FUNCTION_BLOCK basicUVTrojan (* Logica do sistema UV Trojan UV3000Plus (monitoracao Modbus TCP) *)
  (* Standard: 61499-2 *)
  (* Version 1.0, 19/10/2026, Hidryco, Hidryco, 1.0: leitura 41001-41008, canais 1 e 2 (41021-41037, 41061-41077), limpeza 41181-41191; heartbeat 40006 b1 e vigia do heartbeat do SCC *)
  PACKAGE Hidryco.HidrycoLib;
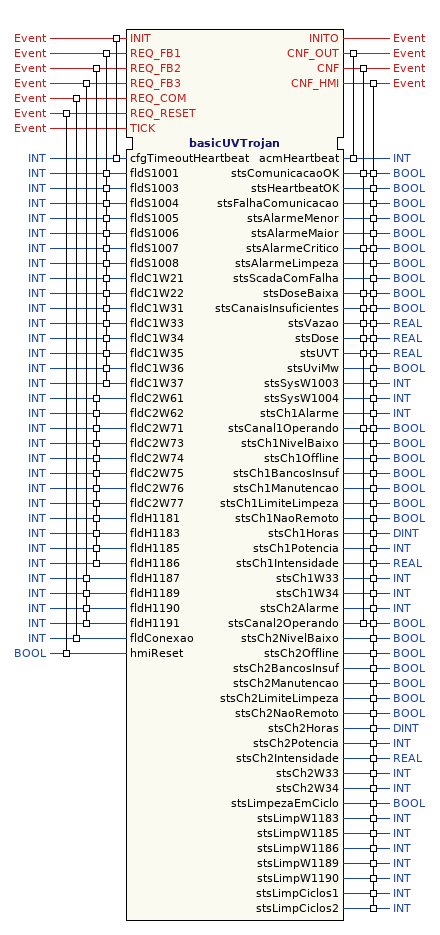
  EVENT_INPUT
    INIT WITH cfgTimeoutHeartbeat; (* Inicializacao *)
    REQ_FB1 WITH fldS1001, fldS1003, fldS1004, fldS1005, fldS1006, fldS1007, fldS1008, fldC1W21, fldC1W22, fldC1W31, fldC1W33, fldC1W34, fldC1W35, fldC1W36, fldC1W37; (* Leitura: sistema e canal 1 *)
    REQ_FB2 WITH fldC2W61, fldC2W62, fldC2W71, fldC2W73, fldC2W74, fldC2W75, fldC2W76, fldC2W77, fldH1181, fldH1183, fldH1185, fldH1186; (* Leitura: canal 2 e limpeza *)
    REQ_FB3 WITH fldH1187, fldH1189, fldH1190, fldH1191; (* Leitura: limpeza (continuacao) *)
    REQ_COM WITH fldConexao; (* Status da conexao Modbus (connStatusInt) *)
    REQ_RESET WITH hmiReset; (* IHM: reconhecimento *)
    TICK; (* Base de tempo de 1 s *)
  END_EVENT
  EVENT_OUTPUT
    INITO; (* Inicializacao concluida *)
    CNF_OUT WITH acmHeartbeat; (* Escrita do heartbeat (40006) *)
    CNF WITH stsComunicacaoOK, stsAlarmeCritico, stsCanal1Operando, stsCanal2Operando, stsCanaisInsuficientes, stsDoseBaixa, stsVazao, stsDose, stsUVT; (* Status para o processo *)
    CNF_HMI WITH stsComunicacaoOK, stsHeartbeatOK, stsFalhaComunicacao, stsAlarmeMenor, stsAlarmeMaior, stsAlarmeCritico, stsAlarmeLimpeza, stsScadaComFalha, stsDoseBaixa, stsCanaisInsuficientes, stsVazao, stsDose, stsUVT, stsUviMw, stsSysW1003, stsSysW1004, stsCh1Alarme, stsCanal1Operando, stsCh1NivelBaixo, stsCh1Offline, stsCh1BancosInsuf, stsCh1Manutencao, stsCh1LimiteLimpeza, stsCh1NaoRemoto, stsCh1Horas, stsCh1Potencia, stsCh1Intensidade, stsCh1W33, stsCh1W34, stsCh2Alarme, stsCanal2Operando, stsCh2NivelBaixo, stsCh2Offline, stsCh2BancosInsuf, stsCh2Manutencao, stsCh2LimiteLimpeza, stsCh2NaoRemoto, stsCh2Horas, stsCh2Potencia, stsCh2Intensidade, stsCh2W33, stsCh2W34, stsLimpezaEmCiclo, stsLimpW1183, stsLimpW1185, stsLimpW1186, stsLimpW1189, stsLimpW1190, stsLimpCiclos1, stsLimpCiclos2; (* Status para a IHM e alarmes *)
  END_EVENT
  VAR_INPUT
    cfgTimeoutHeartbeat : INT := 10; (* Tempo sem alternar o heartbeat do SCC para falha de comunicacao (s) *)
    fldS1001 : INT; (* Registro 41001: alarmes comuns, unidade UVI, heartbeat do SCC *)
    fldS1003 : INT; (* Registro 41003: falhas de sistema 1 *)
    fldS1004 : INT; (* Registro 41004: falhas de sistema 2 *)
    fldS1005 : INT; (* Registro 41005: vazao do sistema *)
    fldS1006 : INT; (* Registro 41006: RED x100 *)
    fldS1007 : INT; (* Registro 41007: UVT x10 *)
    fldS1008 : INT; (* Registro 41008: fator de escala da vazao *)
    fldC1W21 : INT; (* Registro 41021: canal 1 status *)
    fldC1W22 : INT; (* Registro 41022: canal 1 status 2 *)
    fldC1W31 : INT; (* Registro 41031: banco 1A status *)
    fldC1W33 : INT; (* Registro 41033: banco 1A falhas 1 *)
    fldC1W34 : INT; (* Registro 41034: banco 1A falhas 2 *)
    fldC1W35 : INT; (* Registro 41035: banco 1A horas *)
    fldC1W36 : INT; (* Registro 41036: banco 1A potencia *)
    fldC1W37 : INT; (* Registro 41037: banco 1A intensidade x10 *)
    fldC2W61 : INT; (* Registro 41061: canal 2 status *)
    fldC2W62 : INT; (* Registro 41062: canal 2 status 2 *)
    fldC2W71 : INT; (* Registro 41071: banco 2A status *)
    fldC2W73 : INT; (* Registro 41073: banco 2A falhas 1 *)
    fldC2W74 : INT; (* Registro 41074: banco 2A falhas 2 *)
    fldC2W75 : INT; (* Registro 41075: banco 2A horas *)
    fldC2W76 : INT; (* Registro 41076: banco 2A potencia *)
    fldC2W77 : INT; (* Registro 41077: banco 2A intensidade x10 *)
    fldH1181 : INT; (* Registro 41181: limpeza status *)
    fldH1183 : INT; (* Registro 41183: limpeza falhas *)
    fldH1185 : INT; (* Registro 41185: limpeza grupo 1 status *)
    fldH1186 : INT; (* Registro 41186: limpeza grupo 1 falhas *)
    fldH1187 : INT; (* Registro 41187: limpeza grupo 1 ciclos *)
    fldH1189 : INT; (* Registro 41189: limpeza grupo 2 status *)
    fldH1190 : INT; (* Registro 41190: limpeza grupo 2 falhas *)
    fldH1191 : INT; (* Registro 41191: limpeza grupo 2 ciclos *)
    fldConexao : INT; (* connStatusInt (1 = online) *)
    hmiReset : BOOL; (* IHM: reconhecimento *)
  END_VAR
  VAR_OUTPUT
    acmHeartbeat : INT; (* Registro 40006: bit 1 alterna a cada 2 s (heartbeat para o SCC) *)
    stsComunicacaoOK : BOOL; (* Comunicacao Modbus e heartbeat do SCC OK *)
    stsHeartbeatOK : BOOL; (* Heartbeat do SCC (41001.8) alternando *)
    stsFalhaComunicacao : BOOL; (* Falha de comunicacao com o SCC *)
    stsAlarmeMenor : BOOL; (* Alarme comum menor (41001.0) *)
    stsAlarmeMaior : BOOL; (* Alarme comum maior (41001.1) *)
    stsAlarmeCritico : BOOL; (* Alarme comum critico (41001.2) *)
    stsAlarmeLimpeza : BOOL; (* Alarme do sistema de limpeza (41001.3) *)
    stsScadaComFalha : BOOL; (* SCC sem o heartbeat do CLP (41004.4) *)
    stsDoseBaixa : BOOL; (* Dose abaixo do alvo (41003.0) *)
    stsCanaisInsuficientes : BOOL; (* Canais saudaveis insuficientes (41003.1) *)
    stsVazao : REAL; (* Vazao do sistema no SCC (41005 x fator 41008) *)
    stsDose : REAL; (* Dose equivalente RED (mJ/cm2) *)
    stsUVT : REAL; (* Transmitancia UV (%) *)
    stsUviMw : BOOL; (* Unidade da intensidade: FALSE = %, TRUE = mW/cm2 *)
    stsSysW1003 : INT; (* Registro 41003 (diagnostico) *)
    stsSysW1004 : INT; (* Registro 41004 (diagnostico) *)
    stsCh1Alarme : INT; (* Canal 1: 0 normal, 1 menor, 2 maior, 3 critico *)
    stsCanal1Operando : BOOL; (* Canal 1 em operacao *)
    stsCh1NivelBaixo : BOOL; (* Canal 1 nivel de agua baixo *)
    stsCh1Offline : BOOL; (* Canal 1 em modo offline *)
    stsCh1BancosInsuf : BOOL; (* Canal 1 bancos saudaveis insuficientes *)
    stsCh1Manutencao : BOOL; (* Canal 1 em manutencao *)
    stsCh1LimiteLimpeza : BOOL; (* Canal 1 vazao acima do limite de limpeza *)
    stsCh1NaoRemoto : BOOL; (* Banco do canal 1 fora de remoto automatico *)
    stsCh1Horas : DINT; (* Banco do canal 1: horas das lampadas *)
    stsCh1Potencia : INT; (* Banco do canal 1: potencia (%) *)
    stsCh1Intensidade : REAL; (* Banco do canal 1: intensidade UV *)
    stsCh1W33 : INT; (* Banco do canal 1: falhas 1 (diagnostico) *)
    stsCh1W34 : INT; (* Banco do canal 1: falhas 2 (diagnostico) *)
    stsCh2Alarme : INT; (* Canal 2: 0 normal, 1 menor, 2 maior, 3 critico *)
    stsCanal2Operando : BOOL; (* Canal 2 em operacao *)
    stsCh2NivelBaixo : BOOL; (* Canal 2 nivel de agua baixo *)
    stsCh2Offline : BOOL; (* Canal 2 em modo offline *)
    stsCh2BancosInsuf : BOOL; (* Canal 2 bancos saudaveis insuficientes *)
    stsCh2Manutencao : BOOL; (* Canal 2 em manutencao *)
    stsCh2LimiteLimpeza : BOOL; (* Canal 2 vazao acima do limite de limpeza *)
    stsCh2NaoRemoto : BOOL; (* Banco do canal 2 fora de remoto automatico *)
    stsCh2Horas : DINT; (* Banco do canal 2: horas das lampadas *)
    stsCh2Potencia : INT; (* Banco do canal 2: potencia (%) *)
    stsCh2Intensidade : REAL; (* Banco do canal 2: intensidade UV *)
    stsCh2W33 : INT; (* Banco do canal 2: falhas 1 (diagnostico) *)
    stsCh2W34 : INT; (* Banco do canal 2: falhas 2 (diagnostico) *)
    stsLimpezaEmCiclo : BOOL; (* Sistema de limpeza em ciclo *)
    stsLimpW1183 : INT; (* Registro 41183 (diagnostico) *)
    stsLimpW1185 : INT; (* Registro 41185 (diagnostico) *)
    stsLimpW1186 : INT; (* Registro 41186 (diagnostico) *)
    stsLimpW1189 : INT; (* Registro 41189 (diagnostico) *)
    stsLimpW1190 : INT; (* Registro 41190 (diagnostico) *)
    stsLimpCiclos1 : INT; (* Ciclos de limpeza do grupo 1 (canal 1) *)
    stsLimpCiclos2 : INT; (* Ciclos de limpeza do grupo 2 (canal 2) *)
  END_VAR
  VAR
    initDone : BOOL;
    comRecebido : BOOL;
    fb1Recebido : BOOL;
    bComOk : BOOL;
    bHb : BOOL; (* Heartbeat enviado *)
    tHb : INT;
    tHbScc : INT; (* Segundos sem alternar o heartbeat do SCC *)
    bHbScc : BOOL;
    oldHbScc : BOOL;
    lim : INT;
    rFator : REAL;
    w : WORD; (* Palavra em decodificacao *)
    oldHb : INT := -1;
    primeiro : BOOL := TRUE;
    oldAlm : INT := -1; (* Assinatura dos alarmes para disparo imediato *)
    sig : INT;
    oldProc : INT := -1;
  END_VAR
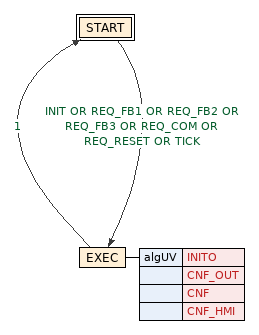
  EC_STATES
    START; (* Estado inicial *)
    EXEC : algUV -> INITO, -> CNF_OUT, -> CNF, -> CNF_HMI; (* Executa a logica; o algoritmo decide quais eventos saem *)
  END_STATES
  EC_TRANSITIONS
    START TO EXEC := INIT OR REQ_FB1 OR REQ_FB2 OR REQ_FB3 OR REQ_COM OR REQ_RESET OR TICK;
    EXEC TO START := 1;
  END_TRANSITIONS
  ALGORITHM algUV IN ST: (* Logica completa do UV (um unico algoritmo) *)
(* =====================================================================
   basicUVTrojan v1.0 - logica do CAT UV_Trojan (HidrycoLib)
   Trojan UV3000Plus, SCC Modicon M580 como servidor Modbus TCP (CP141200010).
   A interface do SCC e somente leitura: o CLP nao liga, nao seleciona canal e
   nao comanda limpeza; so escreve o heartbeat (40006 bit 1, 2 s/2 s). Sem ele
   o SCC acusa SCADA Communication Fault (41004.4).
   Comunicacao OK = conexao Modbus online E heartbeat do SCC (41001.8)
   alternando dentro de cfgTimeoutHeartbeat.
   ===================================================================== *)

INITO   := FALSE;
CNF_OUT := FALSE;
CNF     := FALSE;
CNF_HMI := FALSE;

IF REQ_COM THEN
    comRecebido := TRUE;
END_IF;
IF REQ_FB1 THEN
    fb1Recebido := TRUE;
END_IF;
IF INIT THEN
    initDone := TRUE;
    INITO    := TRUE;
END_IF;
IF NOT initDone THEN
    RETURN;
END_IF;

(* ---- 1. Heartbeat para o SCC e vigia do heartbeat do SCC ---- *)
IF TICK THEN
    tHb := tHb + 1;
    IF tHb >= 2 THEN
        tHb := 0;
        bHb := NOT bHb;
    END_IF;
    IF tHbScc < 32000 THEN
        tHbScc := tHbScc + 1;
    END_IF;
END_IF;
IF bHb THEN
    acmHeartbeat := 2;
ELSE
    acmHeartbeat := 0;
END_IF;
IF (acmHeartbeat <> oldHb) OR primeiro THEN
    CNF_OUT := TRUE;
    oldHb := acmHeartbeat;
END_IF;
w := INT_TO_WORD(fldS1001);
bHbScc := (w AND 16#0100) <> 16#0000;
IF REQ_FB1 AND (bHbScc <> oldHbScc) THEN
    tHbScc := 0;
    oldHbScc := bHbScc;
END_IF;
IF cfgTimeoutHeartbeat > 0 THEN
    lim := cfgTimeoutHeartbeat;
ELSE
    lim := 10;
END_IF;
bComOk := comRecebido AND fb1Recebido AND (fldConexao = 1);
stsHeartbeatOK := bComOk AND (tHbScc < lim);
stsComunicacaoOK := stsHeartbeatOK;
stsFalhaComunicacao := NOT stsComunicacaoOK;

(* ---- 2. Decodificacao (so com comunicacao OK) ---- *)
IF stsComunicacaoOK THEN
    stsAlarmeMenor   := (w AND 16#0001) <> 16#0000;
    stsAlarmeMaior   := (w AND 16#0002) <> 16#0000;
    stsAlarmeCritico := (w AND 16#0004) <> 16#0000;
    stsAlarmeLimpeza := (w AND 16#0008) <> 16#0000;
    stsUviMw         := (w AND 16#0080) <> 16#0000;
    w := INT_TO_WORD(fldS1003);
    stsDoseBaixa := (w AND 16#0001) <> 16#0000;
    stsCanaisInsuficientes := (w AND 16#0002) <> 16#0000;
    w := INT_TO_WORD(fldS1004);
    stsScadaComFalha := (w AND 16#0010) <> 16#0000;
    stsSysW1003 := fldS1003;
    stsSysW1004 := fldS1004;
    CASE fldS1008 OF
        1: rFator := 100.0;
        2: rFator := 10.0;
        4: rFator := 0.1;
        5: rFator := 0.01;
    ELSE
        rFator := 1.0;
    END_CASE;
    stsVazao := INT_TO_REAL(fldS1005) * rFator;
    stsDose  := INT_TO_REAL(fldS1006) / 100.0;
    stsUVT   := INT_TO_REAL(fldS1007) / 10.0;
    (* canal 1 / banco 1A *)
    w := INT_TO_WORD(fldC1W21);
    IF (w AND 16#0004) <> 16#0000 THEN stsCh1Alarme := 3;
    ELSIF (w AND 16#0002) <> 16#0000 THEN stsCh1Alarme := 2;
    ELSIF (w AND 16#0001) <> 16#0000 THEN stsCh1Alarme := 1;
    ELSE stsCh1Alarme := 0;
    END_IF;
    stsCanal1Operando := (w AND 16#0010) <> 16#0000;
    stsCh1NivelBaixo  := (w AND 16#0020) <> 16#0000;
    stsCh1Offline     := (w AND 16#0200) <> 16#0000;
    w := INT_TO_WORD(fldC1W22);
    stsCh1BancosInsuf    := (w AND 16#0002) <> 16#0000;
    stsCh1LimiteLimpeza  := (w AND 16#0020) <> 16#0000;
    stsCh1Manutencao     := (w AND 16#8000) <> 16#0000;
    w := INT_TO_WORD(fldC1W34);
    stsCh1NaoRemoto := (w AND 16#0002) <> 16#0000;
    stsCh1W33 := fldC1W33;
    stsCh1W34 := fldC1W34;
    IF fldC1W35 < 0 THEN stsCh1Horas := INT_TO_DINT(fldC1W35) + 65536; ELSE stsCh1Horas := INT_TO_DINT(fldC1W35); END_IF;
    stsCh1Potencia := fldC1W36;
    stsCh1Intensidade := INT_TO_REAL(fldC1W37) / 10.0;
    (* canal 2 / banco 2A *)
    w := INT_TO_WORD(fldC2W61);
    IF (w AND 16#0004) <> 16#0000 THEN stsCh2Alarme := 3;
    ELSIF (w AND 16#0002) <> 16#0000 THEN stsCh2Alarme := 2;
    ELSIF (w AND 16#0001) <> 16#0000 THEN stsCh2Alarme := 1;
    ELSE stsCh2Alarme := 0;
    END_IF;
    stsCanal2Operando := (w AND 16#0010) <> 16#0000;
    stsCh2NivelBaixo  := (w AND 16#0020) <> 16#0000;
    stsCh2Offline     := (w AND 16#0200) <> 16#0000;
    w := INT_TO_WORD(fldC2W62);
    stsCh2BancosInsuf    := (w AND 16#0002) <> 16#0000;
    stsCh2LimiteLimpeza  := (w AND 16#0020) <> 16#0000;
    stsCh2Manutencao     := (w AND 16#8000) <> 16#0000;
    w := INT_TO_WORD(fldC2W74);
    stsCh2NaoRemoto := (w AND 16#0002) <> 16#0000;
    stsCh2W33 := fldC2W73;
    stsCh2W34 := fldC2W74;
    IF fldC2W75 < 0 THEN stsCh2Horas := INT_TO_DINT(fldC2W75) + 65536; ELSE stsCh2Horas := INT_TO_DINT(fldC2W75); END_IF;
    stsCh2Potencia := fldC2W76;
    stsCh2Intensidade := INT_TO_REAL(fldC2W77) / 10.0;
    (* limpeza (HSC1) *)
    w := INT_TO_WORD(fldH1181);
    stsLimpezaEmCiclo := (w AND 16#0004) <> 16#0000;
    stsLimpW1183 := fldH1183;
    stsLimpW1185 := fldH1185;
    stsLimpW1186 := fldH1186;
    stsLimpW1189 := fldH1189;
    stsLimpW1190 := fldH1190;
    stsLimpCiclos1 := fldH1187;
    stsLimpCiclos2 := fldH1191;
ELSE
    stsAlarmeMenor := FALSE; stsAlarmeMaior := FALSE; stsAlarmeCritico := FALSE; stsAlarmeLimpeza := FALSE;
    stsDoseBaixa := FALSE; stsCanaisInsuficientes := FALSE; stsScadaComFalha := FALSE;
    stsCh1Alarme := 0; stsCanal1Operando := FALSE; stsCh1NivelBaixo := FALSE; stsCh1Offline := FALSE;
    stsCh1BancosInsuf := FALSE; stsCh1Manutencao := FALSE; stsCh1LimiteLimpeza := FALSE; stsCh1NaoRemoto := FALSE;
    stsCh2Alarme := 0; stsCanal2Operando := FALSE; stsCh2NivelBaixo := FALSE; stsCh2Offline := FALSE;
    stsCh2BancosInsuf := FALSE; stsCh2Manutencao := FALSE; stsCh2LimiteLimpeza := FALSE; stsCh2NaoRemoto := FALSE;
    stsLimpezaEmCiclo := FALSE;
END_IF;

(* ---- 3. Eventos: alarmes e estados na hora; valores a cada 1 s ---- *)
sig := 0;
IF stsFalhaComunicacao THEN sig := sig + 1; END_IF;
IF stsAlarmeMenor THEN sig := sig + 2; END_IF;
IF stsAlarmeMaior THEN sig := sig + 4; END_IF;
IF stsAlarmeCritico THEN sig := sig + 8; END_IF;
IF stsAlarmeLimpeza THEN sig := sig + 16; END_IF;
IF stsCanal1Operando THEN sig := sig + 32; END_IF;
IF stsCanal2Operando THEN sig := sig + 64; END_IF;
IF stsCanaisInsuficientes THEN sig := sig + 128; END_IF;
IF stsDoseBaixa THEN sig := sig + 256; END_IF;
IF primeiro OR TICK OR REQ_RESET OR (sig <> oldAlm) THEN
    CNF_HMI := TRUE;
END_IF;
IF primeiro OR TICK OR (sig <> oldAlm) THEN
    CNF := TRUE;
END_IF;
oldAlm := sig;
primeiro := FALSE;
  END_ALGORITHM
END_FUNCTION_BLOCK
